{attribute 'qualified_only'}
{attribute 'strict'}
TYPE E_PistonDefault_CMD :
(
	Close := 0,
	Open,
	Sensors, 		//by actual sensors state
	SensorsClose,	//by actual sensors state, if state wrong close
	SensorsOpen		//by actual sensors state, if state wrong open
);
END_TYPE

(* stored: Version 1.1.0.1, ProductVersion 3.1.4024.12
   DUT E_PistonDefault_CMD: Id {deb4db7c-6913-48ec-9f69-222fb23f7f9a} *)
